// TIA Portal V20 export
// export: Created 2026-11-08T12:24:02.8396068Z, ExportSetting None, DisplayName Totally Integrated Automation Portal, DisplayVersion V20, DisplayName TIA Portal Openness, DisplayVersion V20, DisplayName TIA Portal Version Control Interface, DisplayVersion V20, DisplayName SINAMICS Startdrive Advanced, DisplayVersion V20, DisplayName SINAMICS Startdrive G130, G150, S120, S150, SINAMICS MV, G220, S200, S210, DisplayVersion V20, DisplayName SINAMICS Startdrive G110M, G120, G120C, G120D, G120P, G115D, DisplayVersion V20, DisplayName STEP 7 Professional, DisplayVersion V20, DisplayName STEP 7 Safety, DisplayVersion V20, DisplayName WinCC Basic/Comfort/Advanced, DisplayVersion V20, DisplayName WinCC Unified, DisplayVersion V20
ORGANIZATION_BLOCK "Main"   // OB1, LAD, ProgramCycle
TITLE = "Main Program Sweep (Cycle)"
{ S7_Optimized_Access := 'TRUE' }
// stored: SetENOAutomatically false
   VAR_INPUT
      Initial_Call : Bool;
      Remanence : Bool;
   END_VAR
BEGIN

REGION Network 1
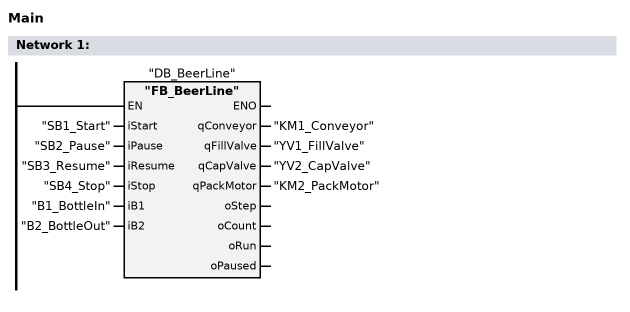
   RUNG wire#powerrail
      "DB_BeerLine"(iStart := "SB1_Start", iPause := "SB2_Pause", iResume := "SB3_Resume", iStop := "SB4_Stop", iB1 := "B1_BottleIn", iB2 := "B2_BottleOut", qConveyor => "KM1_Conveyor", qFillValve => "YV1_FillValve", qCapValve => "YV2_CapValve", qPackMotor => "KM2_PackMotor", oStep =>, oCount =>, oRun =>, oPaused =>)
   END_RUNG
   // the same network as SCL:
   "DB_BeerLine"(iStart := "SB1_Start",   // "FB_BeerLine"
                 iPause := "SB2_Pause",
                 iResume := "SB3_Resume",
                 iStop := "SB4_Stop",
                 iB1 := "B1_BottleIn",
                 iB2 := "B2_BottleOut",
                 qConveyor => "KM1_Conveyor",
                 qFillValve => "YV1_FillValve",
                 qCapValve => "YV2_CapValve",
                 qPackMotor => "KM2_PackMotor");
END_REGION
END_ORGANIZATION_BLOCK
